{attribute 'qualified_only'}
VAR_GLOBAL
    Tank1 : ST_TankHMI;
END_VAR

(* stored: Version 1.1.0.1
   GVL GVL_HMI: Id {c7b210ab-a444-40a9-a550-3710b73030bc} *)
